FUNCTION F_WordToRange_1 : REAL
VAR_INPUT
	wWord 					:WORD;
	rLowLimit 				:REAL;
	rHighLimit 				:REAL;
END_VAR
VAR
END_VAR


F_WordToRange := (rHighLimit - rLowLimit) * WORD_TO_REAL(wWord) * 0.00001525902189669640 + rLowLimit;

END_FUNCTION

(* stored: Version 1.1.0.1, ProductVersion 3.1.4024.15
   POU F_WordToRange_1: Id {bbb638bf-2ed2-4bdf-a595-064b38c8fbca}, SpecialFunc None *)
